Fanuc KAREL source: KT00201.KL

PROGRAM KT00201
%NOLOCKGROUP
VAR
  I1: INTEGER
  B2: BOOLEAN
  OUT: BOOLEAN
BEGIN
  I1 = 2
    B2 = FALSE
  OUT = I1 AND B2
END KT00201
